(* PLC project TBEN_L5_PLC11.project, CODESYS CODESYS V3.5 SP21 Patch 1 *)
(* stored: creationDateTime 2026-11-07T15:35:07.8870036, modificationDateTime 2026-11-07T15:09:07.4034196 *)

// Đọc 4 byte big-endian thành DWORD
FUNCTION F_IolGetU32BE : DWORD
VAR_INPUT
    pBuf  : POINTER TO BYTE;
    uiOff : UINT;
END_VAR

            IF pBuf = 0 THEN
    F_IolGetU32BE := 0;
    RETURN;
END_IF
F_IolGetU32BE := SHL(UINT_TO_DWORD(F_IolGetU16BE(pBuf, uiOff)), 16) OR UINT_TO_DWORD(F_IolGetU16BE(pBuf, uiOff + 2));

          
END_FUNCTION
